(* IEC 61131-3 sources: plcfuzz/testcases/matiec/legacy, 3 files *)

(* ---- boolean_interlock.st ---- *)
PROGRAM BooleanInterlock
  VAR
    StartButton AT %IX0.0 : BOOL;
    StopButton AT %IX0.1 : BOOL;
    MotorEnabled AT %QX0.0 : BOOL;
  END_VAR

  MotorEnabled := StartButton AND NOT StopButton;
END_PROGRAM

CONFIGURATION Config0
  RESOURCE Res0 ON PLC
    TASK MainTask(INTERVAL := T#50ms, PRIORITY := 0);
    PROGRAM Instance0 WITH MainTask : BooleanInterlock;
  END_RESOURCE
END_CONFIGURATION

(* ---- state_machine.st ---- *)
TYPE
  MachineState : (Idle, Starting, Running, Fault) := Idle;
END_TYPE

PROGRAM StateMachine
  VAR
    CurrentState : MachineState := Idle;
  END_VAR
  VAR
    StartButton AT %IX0.0 : BOOL;
    StopButton AT %IX0.1 : BOOL;
    FaultSignal AT %IX0.2 : BOOL;
    RunningLamp AT %QX0.0 : BOOL;
    FaultLamp AT %QX0.1 : BOOL;
  END_VAR

  CASE CurrentState OF
    Idle:
      IF StartButton THEN
        CurrentState := Starting;
      END_IF;
    Starting:
      IF FaultSignal THEN
        CurrentState := Fault;
      ELSE
        CurrentState := Running;
      END_IF;
    Running:
      IF FaultSignal THEN
        CurrentState := Fault;
      ELSIF StopButton THEN
        CurrentState := Idle;
      END_IF;
    Fault:
      IF NOT FaultSignal THEN
        CurrentState := Idle;
      END_IF;
  END_CASE;

  RunningLamp := CurrentState = Running;
  FaultLamp := CurrentState = Fault;
END_PROGRAM

CONFIGURATION Config0
  RESOURCE Res0 ON PLC
    TASK MainTask(INTERVAL := T#50ms, PRIORITY := 0);
    PROGRAM Instance0 WITH MainTask : StateMachine;
  END_RESOURCE
END_CONFIGURATION

(* ---- timer_counter.st ---- *)
PROGRAM TimerCounter
  VAR
    Timer : TON;
    Counter : CTU := (PV := 10);
  END_VAR
  VAR
    Enable AT %IX0.0 : BOOL;
    Reset AT %IX0.1 : BOOL;
    Pulse AT %QX0.0 : BOOL;
  END_VAR

  Timer(IN := Enable, PT := T#500ms);
  Counter(CU := Timer.Q, R := Reset);
  Pulse := Counter.Q;
END_PROGRAM

CONFIGURATION Config0
  RESOURCE Res0 ON PLC
    TASK MainTask(INTERVAL := T#50ms, PRIORITY := 0);
    PROGRAM Instance0 WITH MainTask : TimerCounter;
  END_RESOURCE
END_CONFIGURATION
